{attribute 'qualified_only'}
VAR_GLOBAL PERSISTENT
	
	arrRecipeMarinade	: ARRAY[1..cMax_Prod_Recipe] OF ST_Prod_Recipe;
	arrRecipeColor		: ARRAY[1..cMax_Prod_Recipe] OF ST_Prod_Recipe;
	
	iUserSelected_Marinade	: INT;
	iUserSelected_Color		: INT;
	
	fbProdRecipe_Manage	: FB_ProdRecipe_Manage;
	
	listRecipe_Marinade	: ARRAY[1..cMax_Prod_Recipe] OF STRING(30);
	listRecipe_Color	: ARRAY[1..cMax_Prod_Recipe] OF STRING(30);
	
	dtProdTimePicker	: DATE_AND_TIME;
	dtProdTimeMin		: DATE_AND_TIME;
	dtProdTimeMax		: DATE_AND_TIME;



END_VAR
VAR_GLOBAL CONSTANT 
	cMax_Prod_Recipe	: INT:=10;
	cMaxCompInProduct	: USINT:= 10;
END_VAR

(* stored: Version 1.1.0.1, ProductVersion 3.1.4024.15
   GVL g_Prod: Id {502e9ae9-c438-4303-9edf-0246b0263978} *)
